Fanuc KAREL source: kb00188.compact.KL

PROGRAM KB00188
%STACKSIZE=65535
%PRIORITY=65535
%NOLOCKGROUP
VAR
P1 : STRING[80]
RESULT : INTEGER
BEGIN
P1='A'
RESULT=STR_LEN(P1)
END KB00188
